// TIA Portal V20 export
Screen "200RobotCollision"  1276x673
  ScreenItem "Graphic view_13" at 324,99 size 634x531  Type=HmiGraphicView
  ScreenItem "矩形_6" at -3,69 size 1274x597  Type=HmiRectangle
  ScreenItem "Title_ScreenOverview_X390_Y2" at 438,5 size 551x57  Type=HmiTextBox
  ScreenItem "Line_Header_X0_Y64" at 0,64 size 1274x1  Type=HmiLine
  ScreenItem "permanentareaborderrectangle" at 0,0 size 0x0  Type=HmiRectangle
  ScreenItem "Button_Back" at 2,2 size 90x60  Type=HmiButton
  ScreenItem "Text_3" at 807,91 size 84x39  Type=HmiText
  ScreenItem "Text_4" at 822,617 size 84x39  Type=HmiText
  ScreenItem "Text_5" at 648,611 size 84x39  Type=HmiText
  ScreenItem "Text_6" at 398,91 size 84x39  Type=HmiText
  ScreenItem "Text_18" at 744,583 size 84x73  Type=HmiText
  ScreenItem "Graphic view_6" at 746,-206 size 60x30  Type=HmiGraphicView
  ScreenItem "Graphic view_7" at 746,-594 size 60x30  Type=HmiGraphicView
  ScreenItem "Graphic view_8" at 746,-982 size 60x30  Type=HmiGraphicView
  ScreenItem "Rectangle_5" at 1002,120 size 164x112  Type=HmiRectangle
  ScreenItem "Text_71" at 994,115 size 174x35  Type=HmiText
  ScreenItem "Text_72" at 1025,141 size 123x35  Type=HmiText
  ScreenItem "Text_73" at 1039,169 size 88x35  Type=HmiText
  ScreenItem "Text_74" at 1031,197 size 136x35  Type=HmiText
  ScreenItem "矩形_44" at 1015,204 size 17x17  Type=HmiRectangle
  ScreenItem "矩形_45" at 1015,177 size 17x17  Type=HmiRectangle
  ScreenItem "矩形_46" at 1015,150 size 17x17  Type=HmiRectangle
  ScreenItem "Rectangle_6" at 1006,411 size 164x222  Type=HmiRectangle
  ScreenItem "Text_75" at 998,406 size 174x35  Type=HmiText
  ScreenItem "Text_76" at 1029,432 size 123x35  Type=HmiText
  ScreenItem "Text_77" at 1043,460 size 88x35  Type=HmiText
  ScreenItem "Text_78" at 1035,488 size 136x35  Type=HmiText
  ScreenItem "矩形_47" at 1019,495 size 17x17  Type=HmiRectangle
  ScreenItem "矩形_48" at 1019,468 size 17x17  Type=HmiRectangle
  ScreenItem "矩形_49" at 1019,441 size 17x17  Type=HmiRectangle
  ScreenItem "Text_83" at 1029,542 size 123x35  Type=HmiText
  ScreenItem "Text_84" at 998,516 size 174x35  Type=HmiText
  ScreenItem "矩形_53" at 1019,551 size 17x17  Type=HmiRectangle
  ScreenItem "矩形_54" at 1019,578 size 17x17  Type=HmiRectangle
  ScreenItem "矩形_55" at 1019,605 size 17x17  Type=HmiRectangle
  ScreenItem "Text_85" at 1035,598 size 136x35  Type=HmiText
  ScreenItem "Text_86" at 1043,570 size 88x35  Type=HmiText
  ScreenItem "Graphic view_2" at 749,581 size 60x30  Type=HmiGraphicView
  ScreenItem "Graphic view_4" at 749,545 size 60x30  Type=HmiGraphicView
  ScreenItem "Text_1" at 734,503 size 84x73  Type=HmiText
  ScreenItem "Graphic view_11" at 88,0 size 410x35  Type=HmiGraphicView
  ScreenItem "Graphic view_12" at 0,7 size 410x35  Type=HmiGraphicView
  ScreenItem "Text_2" at 891,492 size 84x73  Type=HmiText
  ScreenItem "Text_9" at 722,202 size 84x73  Type=HmiText
  ScreenItem "Graphic view_1" at 101,0 size 472x35  Type=HmiGraphicView
  ScreenItem "Graphic view_3" at 0,7 size 472x35  Type=HmiGraphicView
  ScreenItem "Text_7" at 296,202 size 84x73  Type=HmiText
  ScreenItem "Text_8" at 580,475 size 84x73  Type=HmiText
  ScreenItem "Rectangle_1" at 179,406 size 164x222  Type=HmiRectangle
  ScreenItem "Text_10" at 171,401 size 174x35  Type=HmiText
  ScreenItem "Text_11" at 202,427 size 123x35  Type=HmiText
  ScreenItem "Text_12" at 216,455 size 88x35  Type=HmiText
  ScreenItem "Text_13" at 208,483 size 136x35  Type=HmiText
  ScreenItem "矩形_1" at 192,490 size 17x17  Type=HmiRectangle
  ScreenItem "矩形_2" at 192,463 size 17x17  Type=HmiRectangle
  ScreenItem "矩形_3" at 192,436 size 17x17  Type=HmiRectangle
  ScreenItem "Text_14" at 202,537 size 123x35  Type=HmiText
  ScreenItem "Text_15" at 171,511 size 174x35  Type=HmiText
  ScreenItem "矩形_4" at 192,546 size 17x17  Type=HmiRectangle
  ScreenItem "矩形_5" at 192,573 size 17x17  Type=HmiRectangle
  ScreenItem "矩形_7" at 192,600 size 17x17  Type=HmiRectangle
  ScreenItem "Text_16" at 208,593 size 136x35  Type=HmiText
  ScreenItem "Text_17" at 216,565 size 88x35  Type=HmiText
  ScreenItem "Rectangle_2" at 176,98 size 164x112  Type=HmiRectangle
  ScreenItem "Text_19" at 168,93 size 174x35  Type=HmiText
  ScreenItem "Text_20" at 199,119 size 123x35  Type=HmiText
  ScreenItem "Text_21" at 213,147 size 88x35  Type=HmiText
  ScreenItem "Text_22" at 205,175 size 136x35  Type=HmiText
  ScreenItem "矩形_8" at 189,182 size 17x17  Type=HmiRectangle
  ScreenItem "矩形_9" at 189,155 size 17x17  Type=HmiRectangle
  ScreenItem "矩形_10" at 189,128 size 17x17  Type=HmiRectangle
